{attribute 'qualified_only'}
VAR_GLOBAL
bEmergencyStop:BOOL;
  nCycleCount : UDINT; // cycles
aMotors:ARRAY [1..3] OF ST_MotorData;
END_VAR
VAR_GLOBAL CONSTANT
cMaxMotors:INT:=3;
END_VAR

(* stored: Version 1.1.0.1
   GVL GVL_Main: Id {9768e80d-482f-4e52-b3ac-9468449bc778} *)
